// TIA Portal V20 export
// export: Created 2026-10-19T18:36:34.9765489Z, ExportSetting WithDefaults, DisplayName Totally Integrated Automation Portal, DisplayVersion V20 Update 6, DisplayName TIA Portal Openness, DisplayVersion V20 Update 6, DisplayName TIA Portal Version Control Interface, DisplayVersion V20 Update 6, DisplayName SINAMICS Startdrive Advanced, DisplayVersion V20 SP1, DisplayName SINAMICS Startdrive G130, G150, S120, S150, SINAMICS MV, G220, S200, S210, DisplayVersion V20 SP1, DisplayName SINAMICS Startdrive G110M, G120, G120C, G120D, G120P, G115D, DisplayVersion V20 SP1, DisplayName STEP 7 Professional, DisplayVersion V20 Update 6, DisplayName STEP 7 Safety, DisplayVersion V20 Update 2, DisplayName WinCC Basic/Comfort/Advanced, DisplayVersion V20 Update 6, DisplayName WinCC Unified, DisplayVersion V20 Update 6
FUNCTION "CNV_Selector_1" : Void   // FC60, SCL
{ S7_Optimized_Access := 'TRUE' }
VERSION : 0.1
// stored: AutoNumber true, IsIECCheckEnabled false, SetENOAutomatically false, UDAEnableTagReadback false
   VAR_INPUT
      Sys_No : UInt;
      Zone : UInt;
      CNV1_2_Selected : UInt;
   END_VAR
   VAR_OUTPUT
      ID : DInt;
      "ID(1)" : DInt;
   END_VAR
BEGIN
   //CNV SCREEN SELECTION
   CASE #Sys_No OF
       0:
           #ID := 0;
           #"ID(1)" := 0;

       1://SYSTEM 1
           CASE #Zone OF
               12: //LEVEL 2
                   "CNV_ID_HMI(1)" := "Settings_DB".LCnv_Sys[#Sys_No].Cnv_Level[#Zone MOD 10].Cnv1.ID; //CNV 1
                   IF "CVTD_CNV2_Selected" = 1 THEN
                       "CNV_ID_HMI" := "Settings_DB".ECnv_Sys[#Sys_No].ID; // EXTRACTOR CONVEYOR
                   ELSIF "CVTD_CNV2_Selected" = 2 THEN
                       "CNV_ID_HMI" := "Settings_DB".LCnv_Sys[#Sys_No].Cnv_Level[#Zone MOD 10].Cnv2.ID; //CNV 2
                   END_IF;
               13: //LEVEL 3
                   "CNV_ID_HMI(1)" := "Settings_DB".LCnv_Sys[#Sys_No].Cnv_Level[#Zone MOD 10].Cnv1.ID; //CNV 1
                   IF "CVTD_CNV2_Selected" = 1 THEN
                       "CNV_ID_HMI" := "Settings_DB".ECnv_Sys[#Sys_No].ID; // EXTRACTOR CONVEYOR
                   ELSIF "CVTD_CNV2_Selected" = 2 THEN
                       "CNV_ID_HMI" := "Settings_DB".LCnv_Sys[#Sys_No].Cnv_Level[#Zone MOD 10].Cnv2.ID; //CNV 2
                   END_IF;
               14: //LEVEL 4
                   "CNV_ID_HMI(1)" := "Settings_DB".LCnv_Sys[#Sys_No].Cnv_Level[#Zone MOD 10].Cnv1.ID; //CNV 1
                   IF "CVTD_CNV2_Selected" = 1 THEN
                       "CNV_ID_HMI" := "Settings_DB".ECnv_Sys[#Sys_No].ID; // EXTRACTOR CONVEYOR
                   ELSIF "CVTD_CNV2_Selected" = 2 THEN
                       "CNV_ID_HMI" := "Settings_DB".LCnv_Sys[#Sys_No].Cnv_Level[#Zone MOD 10].Cnv2.ID; //CNV 2
                   END_IF;
               15: //LEVEL 5
                   "CNV_ID_HMI(1)" := "Settings_DB".LCnv_Sys[#Sys_No].Cnv_Level[#Zone MOD 10].Cnv1.ID; //CNV 1
                   IF "CVTD_CNV2_Selected" = 1 THEN
                       "CNV_ID_HMI" := "Settings_DB".ECnv_Sys[#Sys_No].ID; // EXTRACTOR CONVEYOR
                   ELSIF "CVTD_CNV2_Selected" = 2 THEN
                       "CNV_ID_HMI" := "Settings_DB".LCnv_Sys[#Sys_No].Cnv_Level[#Zone MOD 10].Cnv2.ID; //CNV 2
                   END_IF;
               16: //LEVEL 6
                   "CNV_ID_HMI(1)" := "Settings_DB".LCnv_Sys[#Sys_No].Cnv_Level[#Zone MOD 10].Cnv1.ID; //CNV 1
                   IF "CVTD_CNV2_Selected" = 1 THEN
                       "CNV_ID_HMI" := "Settings_DB".ECnv_Sys[#Sys_No].ID; // EXTRACTOR CONVEYOR
                   ELSIF "CVTD_CNV2_Selected" = 2 THEN
                       "CNV_ID_HMI" := "Settings_DB".LCnv_Sys[#Sys_No].Cnv_Level[#Zone MOD 10].Cnv2.ID; //CNV 2
                   END_IF;
           END_CASE;

       2://SYSTEM 2
           CASE #Zone OF
               12: //LEVEL 2
                   "CNV_ID_HMI(1)" := "Settings_DB".LCnv_Sys[#Sys_No].Cnv_Level[#Zone MOD 10].Cnv1.ID; //CNV 1
                   IF "CVTD_CNV2_Selected" = 1 THEN
                       "CNV_ID_HMI" := "Settings_DB".ECnv_Sys[#Sys_No].ID; // EXTRACTOR CONVEYOR
                   ELSIF "CVTD_CNV2_Selected" = 2 THEN
                       "CNV_ID_HMI" := "Settings_DB".LCnv_Sys[#Sys_No].Cnv_Level[#Zone MOD 10].Cnv2.ID; //CNV 2
                   END_IF;
               13: //LEVEL 3
                   "CNV_ID_HMI(1)" := "Settings_DB".LCnv_Sys[#Sys_No].Cnv_Level[#Zone MOD 10].Cnv1.ID; //CNV 1
                   IF "CVTD_CNV2_Selected" = 1 THEN
                       "CNV_ID_HMI" := "Settings_DB".ECnv_Sys[#Sys_No].ID; // EXTRACTOR CONVEYOR
                   ELSIF "CVTD_CNV2_Selected" = 2 THEN
                       "CNV_ID_HMI" := "Settings_DB".LCnv_Sys[#Sys_No].Cnv_Level[#Zone MOD 10].Cnv2.ID; //CNV 2
                   END_IF;
               14: //LEVEL 4
                   "CNV_ID_HMI(1)" := "Settings_DB".LCnv_Sys[#Sys_No].Cnv_Level[#Zone MOD 10].Cnv1.ID; //CNV 1
                   IF "CVTD_CNV2_Selected" = 1 THEN
                       "CNV_ID_HMI" := "Settings_DB".ECnv_Sys[#Sys_No].ID; // EXTRACTOR CONVEYOR
                   ELSIF "CVTD_CNV2_Selected" = 2 THEN
                       "CNV_ID_HMI" := "Settings_DB".LCnv_Sys[#Sys_No].Cnv_Level[#Zone MOD 10].Cnv2.ID; //CNV 2
                   END_IF;
               15: //LEVEL 5
                   "CNV_ID_HMI(1)" := "Settings_DB".LCnv_Sys[#Sys_No].Cnv_Level[#Zone MOD 10].Cnv1.ID; //CNV 1
                   IF "CVTD_CNV2_Selected" = 1 THEN
                       "CNV_ID_HMI" := "Settings_DB".ECnv_Sys[#Sys_No].ID; // EXTRACTOR CONVEYOR
                   ELSIF "CVTD_CNV2_Selected" = 2 THEN
                       "CNV_ID_HMI" := "Settings_DB".LCnv_Sys[#Sys_No].Cnv_Level[#Zone MOD 10].Cnv2.ID; //CNV 2
                   END_IF;
               16: //LEVEL 6
                   "CNV_ID_HMI(1)" := "Settings_DB".LCnv_Sys[#Sys_No].Cnv_Level[#Zone MOD 10].Cnv1.ID; //CNV 1
                   IF "CVTD_CNV2_Selected" = 1 THEN
                       "CNV_ID_HMI" := "Settings_DB".ECnv_Sys[#Sys_No].ID; // EXTRACTOR CONVEYOR
                   ELSIF "CVTD_CNV2_Selected" = 2 THEN
                       "CNV_ID_HMI" := "Settings_DB".LCnv_Sys[#Sys_No].Cnv_Level[#Zone MOD 10].Cnv2.ID; //CNV 2
                   END_IF;
           END_CASE;
   END_CASE;
END_FUNCTION
